ADAPTER AFIFO_UINT (* Adapter fuer FIFO_UINT (FIFO_adapter): Konsument haengt per Socket an - DATA liefert PLUG->SOCKET den naechsten Wert, PROCESSED quittiert SOCKET->PLUG dessen Verarbeitung. Kein eigener Event-Baustein auf Konsumentenseite noetig - der Rueckkanal des Adapters selbst traegt die Quittung. *)
  (* Standard: 61499-1; Description: Copyright (c) 2026 Meisterschulen am Ostbahnhof This program and the accompanying materials are made available under the terms of the Eclipse Public License 2.0 which is available at https://www.eclipse.org/legal/epl-2.0/ SPDX-License-Identifier: EPL-2.0 *)
  (* Version 1.1, 2026-11-08, Franz Höpfinger, Meisterschulen am Ostbahnhof, N (Fuellstand der Queue) wird mit DATA mitgeliefert. *)
  (* Version 1.0, 2026-10-13, Franz Höpfinger, Meisterschulen am Ostbahnhof, initial API and implementation and/or initial documentation *)
  PACKAGE FIFO_adapter;
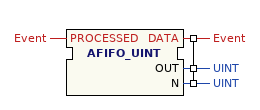
  EVENT_INPUT
    PROCESSED; (* Konsument (SOCKET) bestaetigt: OUT ist verarbeitet, der naechste Wert (falls vorhanden) kann geliefert werden *)
  END_EVENT
  EVENT_OUTPUT
    DATA WITH OUT, N; (* PLUG (FIFO) liefert einen neuen Wert - es folgt kein weiteres DATA, bevor nicht PROCESSED eingetroffen ist *)
  END_EVENT
  VAR_OUTPUT
    OUT : UINT; (* Gelieferter Wert, gueltig bis zur naechsten PROCESSED-Bestaetigung *)
    N : UINT; (* Anzahl der danach noch wartenden Elemente in der Queue *)
  END_VAR
END_ADAPTER
